// TIA Portal V20 export
Screen "200RB04_J5"  1276x673
  ScreenItem "Graphic view_2" at 48,88 size 878x526  Type=HmiGraphicView
  ScreenItem "Line_Header_X0_Y64" at -3,67 size 1276x0  Type=HmiLine
  ScreenItem "permanentareaborderrectangle" at 0,0 size 0x0  Type=HmiRectangle
  ScreenItem "Button_Back" at 2,2 size 90x60  Type=HmiButton
  ScreenItem "文本域_11" at 672,68 size 134x40  Type=HmiTextBox
  ScreenItem "Rectangle_2" at 0,0 size 166x43  Type=HmiRectangle
  ScreenItem "文本域_2" at 2,1 size 134x40  Type=HmiTextBox
  ScreenItem "圆_1" at 0,0 size 100x30  Type=HmiCircle
  ScreenItem "圆_2" at 0,0 size 100x30  Type=HmiCircle
  ScreenItem "Rectangle_3" at 0,0 size 166x43  Type=HmiRectangle
  ScreenItem "文本域_3" at 2,1 size 134x40  Type=HmiTextBox
  ScreenItem "圆_3" at 0,0 size 100x30  Type=HmiCircle
  ScreenItem "圆_4" at 0,0 size 100x30  Type=HmiCircle
  ScreenItem "文本域_1" at 317,160 size 134x40  Type=HmiTextBox
  ScreenItem "文本域_4" at 949,326 size 134x40  Type=HmiTextBox
  ScreenItem "文本域_9" at 950,444 size 134x40  Type=HmiTextBox
  ScreenItem "文本域_13" at 577,578 size 134x40  Type=HmiTextBox
  ScreenItem "文本域_12" at 328,464 size 134x40  Type=HmiTextBox
  ScreenItem "Rectangle_13" at 0,0 size 166x43  Type=HmiRectangle
  ScreenItem "文本域_14" at 2,1 size 134x40  Type=HmiTextBox
  ScreenItem "圆_5" at 0,0 size 100x30  Type=HmiCircle
  ScreenItem "圆_6" at 0,0 size 100x30  Type=HmiCircle
  ScreenItem "Line_2" at 790,284 size 148x3  Type=HmiLine
  ScreenItem "Line_4" at 452,183 size 140x120  Type=HmiLine
  ScreenItem "Line_8" at 704,336 size 244x129  Type=HmiLine
  ScreenItem "Line_9" at 464,417 size 124x70  Type=HmiLine
  ScreenItem "Line_1" at 647,480 size 84x100  Type=HmiLine
  ScreenItem "Rectangle_1" at 0,0 size 52x43  Type=HmiRectangle
  ScreenItem "Title_ScreenOverview_X390_Y2_111" at 0,21 size 25x21  Type=HmiTextBox
  ScreenItem "Title_ScreenOverview_X390_Y2_90" at 27,21 size 25x21  Type=HmiTextBox
  ScreenItem "Title_ScreenOverview_X390_Y2_88" at 0,1 size 52x19  Type=HmiTextBox
  ScreenItem "Rectangle_4" at 0,0 size 52x43  Type=HmiRectangle
  ScreenItem "Title_ScreenOverview_X390_Y2_2" at 0,21 size 25x21  Type=HmiTextBox
  ScreenItem "Title_ScreenOverview_X390_Y2_3" at 27,21 size 25x21  Type=HmiTextBox
  ScreenItem "Title_ScreenOverview_X390_Y2_4" at 0,1 size 52x19  Type=HmiTextBox
  ScreenItem "Title_ScreenOverview_X390_Y2_20" at 713,132 size 25x21  Type=HmiTextBox
  ScreenItem "Rectangle_10" at 713,111 size 52x43  Type=HmiRectangle
  ScreenItem "Title_ScreenOverview_X390_Y2_21" at 740,132 size 25x21  Type=HmiTextBox
  ScreenItem "Title_ScreenOverview_X390_Y2_22" at 713,112 size 52x19  Type=HmiTextBox
  ScreenItem "Title_ScreenOverview_X390_Y2_5" at 393,4 size 510x57  Type=HmiTextBox
  ScreenItem "Line_3" at 454,128 size 136x150  Type=HmiLine
  ScreenItem "Line_5" at 619,87 size 54x50  Type=HmiLine
  ScreenItem "Line_6" at 734,152 size 197x117  Type=HmiLine
  ScreenItem "Line_10" at 660,224 size 276x88  Type=HmiLine
  ScreenItem "Line_11" at 783,331 size 167x18  Type=HmiLine
  ScreenItem "Fusszeile_Button_ManualOPMode1_1" at 1184,2 size 90x60  Type=HmiButton
  ScreenItem "Title_ScreenOverview_X390_Y2_1" at 1138,86 size 139x57  Type=HmiTextBox
  ScreenItem "Title_ScreenOverview_X390_Y2_6" at 1138,152 size 139x57  Type=HmiTextBox
  ScreenItem "Title_ScreenOverview_X390_Y2_7" at 1138,152 size 139x57  Type=HmiTextBox
  ScreenItem "Rectangle_11" at 0,0 size 52x43  Type=HmiRectangle
  ScreenItem "Title_ScreenOverview_X390_Y2_23" at 0,21 size 25x21  Type=HmiTextBox
  ScreenItem "Title_ScreenOverview_X390_Y2_24" at 27,21 size 25x21  Type=HmiTextBox
  ScreenItem "Title_ScreenOverview_X390_Y2_25" at 0,1 size 52x19  Type=HmiTextBox
  ScreenItem "Title_ScreenOverview_X390_Y2_26" at 0,22 size 25x21  Type=HmiTextBox
  ScreenItem "Title_ScreenOverview_X390_Y2_27" at 27,22 size 25x21  Type=HmiTextBox
  ScreenItem "Title_ScreenOverview_X390_Y2_28" at 0,2 size 52x19  Type=HmiTextBox
  ScreenItem "Rectangle_12" at 0,0 size 52x43  Type=HmiRectangle
  ScreenItem "Title_ScreenOverview_X390_Y2_17" at 0,21 size 25x21  Type=HmiTextBox
  ScreenItem "Title_ScreenOverview_X390_Y2_18" at 27,21 size 25x21  Type=HmiTextBox
  ScreenItem "Title_ScreenOverview_X390_Y2_19" at 0,1 size 52x19  Type=HmiTextBox
  ScreenItem "Rectangle_9" at 0,0 size 52x43  Type=HmiRectangle
  ScreenItem "Rectangle_5" at 0,0 size 166x43  Type=HmiRectangle
  ScreenItem "文本域_5" at 2,1 size 134x40  Type=HmiTextBox
  ScreenItem "圆_7" at 0,0 size 100x30  Type=HmiCircle
  ScreenItem "圆_8" at 0,0 size 100x30  Type=HmiCircle
